FUNCTION_BLOCK DS18B20 (* Temperature of a DS18B20 on the 1-Wire bus of logiBUS *)
  (* Standard: 61499-2; Description: Copyright (c) 2026 HR Agrartechnik GmbH This program and the accompanying materials are made available under the terms of the Eclipse Public License 2.0 which is available at https://www.eclipse.org/legal/epl-2.0/ SPDX-License-Identifier: EPL-2.0 The firmware measures all DS18B20 of the bus about once per second (12 bit, 0.0625 °C). Bus GPIO per board (Trainer20: GPIO3); an external 4.7 kOhm pull-up to 3.3 V is recommended. Selection: ROM <> 0 selects the sensor with this ROM code, ROM = 0 the sensor Index in search order (0 = first). ROMO shows the ROM code actually used: write it to ROM to keep the sensor when others are added. IND after each measurement of the sensor and when the state changes. QO = TRUE: Temp is valid. STATUS: OK, no 1-Wire bus, sensor not found, read error, power-on value 85 °C, no value yet. Several DS18B20 FBs may use the same bus (up to 8). *)
  (* Version 1.0, 2026-11-26, Franz Höpfinger, initial API and implementation and/or initial documentation *)
  PACKAGE logiBUS::onewire;
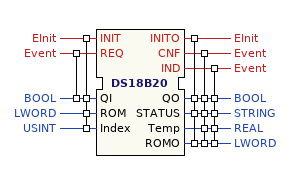
  EVENT_INPUT
    INIT : EInit WITH QI, ROM, Index; (* Service Initialization *)
    REQ WITH QI; (* Read the last value *)
  END_EVENT
  EVENT_OUTPUT
    INITO : EInit WITH QO, STATUS, ROMO; (* Initialization Confirm *)
    CNF WITH QO, STATUS, Temp, ROMO; (* Confirmation of Requested Service *)
    IND WITH QO, STATUS, Temp, ROMO; (* New measurement or changed state *)
  END_EVENT
  VAR_INPUT
    QI : BOOL; (* Event Input Qualifier *)
    ROM : LWORD; (* ROM code of the sensor, 0 = use Index *)
    Index : USINT; (* Sensor in search order (0 = first), if ROM = 0 *)
  END_VAR
  VAR_OUTPUT
    QO : BOOL; (* TRUE: Temp is valid *)
    STATUS : STRING; (* Service Status *)
    Temp : REAL; (* Temperature in °C *)
    ROMO : LWORD; (* ROM code of the sensor used (0 = none) *)
  END_VAR
END_FUNCTION_BLOCK
